(* IEC 61131-3 sources: 2026_Projet_YGO_ExcavatriceDragage/ARCHIVES/Code/PLC_TESTS/BRICKS, 6 files *)

(* ---- FB_TestCheck.st ---- *)
FUNCTION_BLOCK FB_TestCheck
VAR_INPUT
    Config      : ST_TestCheckConfig;
    Evaluate    : BOOL;
END_VAR
VAR_IN_OUT
    ProbeBool   : ARRAY[1..GVL_PLC_Tests_Const.MaxProbeBool] OF BOOL;
    ProbeDint   : ARRAY[1..GVL_PLC_Tests_Const.MaxProbeDint] OF DINT;
    ProbeReal   : ARRAY[1..GVL_PLC_Tests_Const.MaxProbeReal] OF REAL;
END_VAR
VAR_OUTPUT
    Passed       : BOOL;
    Failed       : BOOL;
    Pending      : BOOL;
    FailReason   : E_TestFailReason;
    ObservedBool : BOOL;
    ObservedDint : DINT;
    ObservedReal : REAL;
END_VAR
VAR
    RisingTrig   : R_TRIG;
    FallingTrig  : F_TRIG;
    StableTimer  : TON;
    EvaluateTrig : R_TRIG;
    Cond         : BOOL;
    ProbeIdxLocal : INT;
END_VAR
// === IMPLEMENTATION ===
// Toujours mettre à jour les triggers, avec borne validée AVANT l'accès.
ProbeIdxLocal := Config.ProbeIdx;
IF ProbeIdxLocal >= 1 THEN
    IF ProbeIdxLocal <= GVL_PLC_Tests_Const.MaxProbeBool THEN
        RisingTrig(CLK := ProbeBool[ProbeIdxLocal]);
        FallingTrig(CLK := ProbeBool[ProbeIdxLocal]);
    ELSE
        RisingTrig(CLK := FALSE);
        FallingTrig(CLK := FALSE);
    END_IF;
ELSE
    RisingTrig(CLK := FALSE);
    FallingTrig(CLK := FALSE);
END_IF;

EvaluateTrig(CLK := Evaluate);

IF EvaluateTrig.Q THEN
    Passed := FALSE;
    Failed := FALSE;
    Pending := FALSE;
    FailReason := E_TestFailReason.FAIL_NONE;
    StableTimer(IN := FALSE);
END_IF;

// Mise à jour des valeurs observées
IF Config.ProbeIdx >= 1 THEN
    CASE Config.Kind OF
        E_TestCheckKind.BOOL_EQUAL, E_TestCheckKind.BOOL_RISING, E_TestCheckKind.BOOL_FALLING:
            IF Config.ProbeIdx <= GVL_PLC_Tests_Const.MaxProbeBool THEN
                ObservedBool := ProbeBool[ProbeIdxLocal];
            END_IF;
        E_TestCheckKind.DINT_EQUAL, E_TestCheckKind.DINT_NOT_EQUAL, E_TestCheckKind.DINT_IN_RANGE,
        E_TestCheckKind.WORD_MASK_ALL, E_TestCheckKind.WORD_MASK_ANY, E_TestCheckKind.WORD_MASK_NONE:
            IF Config.ProbeIdx <= GVL_PLC_Tests_Const.MaxProbeDint THEN
                ObservedDint := ProbeDint[ProbeIdxLocal];
            END_IF;
        E_TestCheckKind.REAL_IN_RANGE:
            IF Config.ProbeIdx <= GVL_PLC_Tests_Const.MaxProbeReal THEN
                ObservedReal := ProbeReal[ProbeIdxLocal];
            END_IF;
    END_CASE;
END_IF;

// Évaluation de la condition logique (Cond)
Cond := FALSE;
IF Config.ProbeIdx >= 1 THEN
    CASE Config.Kind OF
        E_TestCheckKind.BOOL_EQUAL:
            IF Config.ProbeIdx <= GVL_PLC_Tests_Const.MaxProbeBool THEN
                Cond := (ObservedBool = Config.ExpectedBool);
            END_IF;

        E_TestCheckKind.BOOL_RISING:
            IF Config.ProbeIdx <= GVL_PLC_Tests_Const.MaxProbeBool THEN
                Cond := RisingTrig.Q;
            END_IF;

        E_TestCheckKind.BOOL_FALLING:
            IF Config.ProbeIdx <= GVL_PLC_Tests_Const.MaxProbeBool THEN
                Cond := FallingTrig.Q;
            END_IF;

        E_TestCheckKind.DINT_EQUAL:
            IF Config.ProbeIdx <= GVL_PLC_Tests_Const.MaxProbeDint THEN
                Cond := (ObservedDint = Config.ExpectedDint);
            END_IF;

        E_TestCheckKind.DINT_NOT_EQUAL:
            IF Config.ProbeIdx <= GVL_PLC_Tests_Const.MaxProbeDint THEN
                Cond := (ObservedDint <> Config.ExpectedDint);
            END_IF;

        E_TestCheckKind.DINT_IN_RANGE:
            IF Config.ProbeIdx <= GVL_PLC_Tests_Const.MaxProbeDint THEN
                Cond := (ObservedDint >= Config.ExpectedMin AND ObservedDint <= Config.ExpectedMax);
            END_IF;

        E_TestCheckKind.WORD_MASK_ALL:
            IF Config.ProbeIdx <= GVL_PLC_Tests_Const.MaxProbeDint THEN
                Cond := ((DINT_TO_WORD(ObservedDint) AND Config.Mask) = Config.Mask);
            END_IF;

        E_TestCheckKind.WORD_MASK_ANY:
            IF Config.ProbeIdx <= GVL_PLC_Tests_Const.MaxProbeDint THEN
                Cond := ((DINT_TO_WORD(ObservedDint) AND Config.Mask) <> 0);
            END_IF;

        E_TestCheckKind.WORD_MASK_NONE:
            IF Config.ProbeIdx <= GVL_PLC_Tests_Const.MaxProbeDint THEN
                Cond := ((DINT_TO_WORD(ObservedDint) AND Config.Mask) = 0);
            END_IF;

        E_TestCheckKind.REAL_IN_RANGE:
            IF Config.ProbeIdx <= GVL_PLC_Tests_Const.MaxProbeReal THEN
                Cond := (ObservedReal >= Config.RealMin AND ObservedReal <= Config.RealMax);
            END_IF;
    END_CASE;
END_IF;

// Application du mode d'évaluation
IF Evaluate THEN
    CASE Config.Mode OF
        E_TestCheckMode.CHECK_INSTANT:
            IF EvaluateTrig.Q THEN
                IF Cond THEN
                    Passed := TRUE;
                    Failed := FALSE;
                    Pending := FALSE;
                ELSE
                    Passed := FALSE;
                    Failed := TRUE;
                    Pending := FALSE;
                    FailReason := E_TestFailReason.FAIL_CHECK;
                END_IF;
            END_IF;

        E_TestCheckMode.CHECK_WAIT_UNTIL:
            IF NOT Passed AND NOT Failed THEN
                StableTimer(IN := Cond, PT := Config.StablePT);
                IF StableTimer.Q THEN
                    Passed := TRUE;
                    Failed := FALSE;
                    Pending := FALSE;
                ELSE
                    Pending := TRUE;
                END_IF;
            END_IF;

        E_TestCheckMode.CHECK_INVARIANT:
            IF NOT Cond THEN
                Passed := FALSE;
                Failed := TRUE;
                Pending := FALSE;
                FailReason := E_TestFailReason.FAIL_INVARIANT;
            ELSE
                Passed := TRUE;
                Failed := FALSE;
                Pending := FALSE;
            END_IF;

        E_TestCheckMode.CHECK_NEVER_DURING:
            IF NOT Failed THEN
                IF Cond THEN
                    Passed := FALSE;
                    Failed := TRUE;
                    Pending := FALSE;
                    FailReason := E_TestFailReason.FAIL_CHECK;
                ELSE
                    Pending := TRUE;
                END_IF;
            END_IF;
    END_CASE;
ELSE
    Passed := FALSE;
    Failed := FALSE;
    Pending := FALSE;
    StableTimer(IN := FALSE);
END_IF;

(* ---- FB_TestEdgeCounter.st ---- *)
FUNCTION_BLOCK FB_TestEdgeCounter
VAR_INPUT
    Arm         : BOOL;
    Signal      : BOOL;
    CountRising : BOOL; // TRUE pour fronts montants, FALSE pour descendants
    ExpectedMin : DINT;
    ExpectedMax : DINT;
END_VAR
VAR_OUTPUT
    Count       : DINT;
    InRange     : BOOL;
END_VAR
VAR
    TrigRising  : R_TRIG;
    TrigFalling : F_TRIG;
END_VAR
// === IMPLEMENTATION ===
TrigRising(CLK := Signal);
TrigFalling(CLK := Signal);

IF NOT Arm THEN
    Count := 0;
    InRange := FALSE;
    RETURN;
END_IF;

IF CountRising AND TrigRising.Q THEN
    Count := Count + 1;
ELSIF NOT CountRising AND TrigFalling.Q THEN
    Count := Count + 1;
END_IF;

InRange := (Count >= ExpectedMin AND Count <= ExpectedMax);

(* ---- FB_TestEventOrder.st ---- *)
FUNCTION_BLOCK FB_TestEventOrder
VAR_INPUT
    Arm       : BOOL;
    EventA    : BOOL;
    EventB    : BOOL;
    TimeoutPT : TIME;
END_VAR
VAR_OUTPUT
    OrderOk   : BOOL;
    Failed    : BOOL;
END_VAR
VAR
    TrigA     : R_TRIG;
    TrigB     : R_TRIG;
    Timer     : TON;
    HasA      : BOOL;
END_VAR
// === IMPLEMENTATION ===
TrigA(CLK := EventA);
TrigB(CLK := EventB);

IF NOT Arm THEN
    OrderOk := FALSE;
    Failed  := FALSE;
    HasA    := FALSE;
    Timer(IN := FALSE);
    RETURN;
END_IF;

// Échec immédiat si B se produit avant A
IF TrigB.Q AND NOT HasA THEN
    Failed  := TRUE;
    OrderOk := FALSE;
END_IF;

// Mémorisation de la survenue de A
IF TrigA.Q AND NOT Failed AND NOT OrderOk THEN
    HasA := TRUE;
END_IF;

// Armement du timeout une fois que A s'est produit
Timer(IN := HasA AND NOT OrderOk AND NOT Failed, PT := TimeoutPT);

IF Timer.Q THEN
    Failed  := TRUE;
    OrderOk := FALSE;
END_IF;

// Validation du succès si B arrive après A et dans les temps
IF HasA AND TrigB.Q AND NOT Failed THEN
    OrderOk := TRUE;
END_IF;

(* ---- FB_TestStimulus.st ---- *)
FUNCTION_BLOCK FB_TestStimulus
VAR_INPUT
    Config     : ST_TestStimAnalogConfig;
    Start      : BOOL;
    Abort      : BOOL;
END_VAR
VAR_OUTPUT
    OutBool    : BOOL;
    OutReal    : REAL;
    OutActive  : BOOL;
    Done       : BOOL;
END_VAR
VAR
    StartTrig   : R_TRIG;
    Timer       : TON;
    SeqTimer    : TON;
    Ramp        : RAMP_REAL;
    ActiveIndex : INT;
    Running     : BOOL;
    Rate        : REAL;
END_VAR
// === IMPLEMENTATION ===
StartTrig(CLK := Start);

// Gestion de l'arrêt ou de l'inactivité
IF Abort OR (NOT Running AND NOT StartTrig.Q) THEN
    Running := FALSE;
    OutActive := FALSE;
    OutBool := FALSE;
    OutReal := 0.0;
    Done := FALSE;
    Timer(IN := FALSE);
    SeqTimer(IN := FALSE);
    Ramp(RESET := TRUE, IN := 0.0);
    RETURN;
END_IF;

// Lancement sur front montant de Start
IF StartTrig.Q THEN
    Running := TRUE;
    Done := FALSE;
    OutActive := TRUE;
    ActiveIndex := 1;
    Timer(IN := FALSE);
    SeqTimer(IN := FALSE);

    CASE Config.Kind OF
        E_TestStimKind.STIM_PULSE_BOOL:
            OutBool := TRUE;
            Timer(IN := TRUE, PT := Config.PulsePT);

        E_TestStimKind.STIM_RAMP_REAL:
            Ramp(RESET := TRUE, IN := Config.StartReal);
            IF Config.RampPT > T#0s THEN
                // Calcul de la vitesse par seconde
                Rate := ABS(Config.TargetReal - Config.StartReal) / (TIME_TO_REAL(Config.RampPT) / 1000.0);
            ELSE
                Rate := ABS(Config.TargetReal - Config.StartReal);
            END_IF;
            Timer(IN := TRUE, PT := Config.RampPT);

        E_TestStimKind.STIM_SEQUENCE_REAL:
            IF Config.SeqCount >= 1 THEN
                OutReal := Config.SeqValues[1];
                SeqTimer(IN := TRUE, PT := Config.SeqDwellPT);
            ELSE
                Running := FALSE;
                OutActive := FALSE;
                Done := TRUE;
            END_IF;
    END_CASE;
END_IF;

// Éxecution logique quand le stimulus tourne
IF Running THEN
    CASE Config.Kind OF
        E_TestStimKind.STIM_PULSE_BOOL:
            Timer();
            IF Timer.Q THEN
                OutBool := FALSE;
                Running := FALSE;
                OutActive := FALSE;
                Done := TRUE;
                Timer(IN := FALSE);
            END_IF;

        E_TestStimKind.STIM_RAMP_REAL:
            Timer();
            Ramp(RESET := FALSE, IN := Config.TargetReal, ASCEND := Rate, DESCEND := Rate, TIMEBASE := T#1s);
            OutReal := Ramp.OUT;
            IF Timer.Q THEN
                OutReal := Config.TargetReal; // Assure la valeur cible exacte à la fin
                Running := FALSE;
                OutActive := FALSE;
                Done := TRUE;
                Timer(IN := FALSE);
            END_IF;

        E_TestStimKind.STIM_SEQUENCE_REAL:
            SeqTimer();
            IF SeqTimer.Q THEN
                SeqTimer(IN := FALSE);
                ActiveIndex := ActiveIndex + 1;
                IF ActiveIndex > Config.SeqCount OR ActiveIndex > GVL_PLC_Tests_Const.MaxSeqValues THEN
                    Running := FALSE;
                    OutActive := FALSE;
                    Done := TRUE;
                ELSE
                    OutReal := Config.SeqValues[ActiveIndex];
                    SeqTimer(IN := TRUE, PT := Config.SeqDwellPT);
                END_IF;
            END_IF;
    END_CASE;
END_IF;

(* ---- FB_TestStopwatch.st ---- *)
FUNCTION_BLOCK FB_TestStopwatch
VAR_INPUT
    Arm             : BOOL;
    StartEvent      : BOOL;
    StopEvent       : BOOL;
    ExpectedMinMs   : DINT;
    ExpectedMaxMs   : DINT;
END_VAR
VAR_OUTPUT
    ElapsedMs       : DINT;
    Done            : BOOL;
    InWindow        : BOOL;
END_VAR
VAR
    StartTrig       : R_TRIG;
    StopTrig        : R_TRIG;
    Running         : BOOL;
    CycleCount      : UDINT;
END_VAR
// === IMPLEMENTATION ===
StartTrig(CLK := StartEvent);
StopTrig(CLK := StopEvent);

IF NOT Arm THEN
    Running := FALSE;
    Done := FALSE;
    InWindow := FALSE;
    ElapsedMs := 0;
    CycleCount := 0;
    RETURN;
END_IF;

IF StartTrig.Q AND NOT Running AND NOT Done THEN
    Running := TRUE;
    CycleCount := 0;
END_IF;

IF Running THEN
    // Incrémente le compteur de cycles
    CycleCount := CycleCount + 1;
    ElapsedMs := UDINT_TO_DINT(CycleCount * INT_TO_UDINT(GVL_PLC_Tests_Const.TaskCycleMs));

    IF StopTrig.Q THEN
        Running := FALSE;
        Done := TRUE;
        InWindow := (ElapsedMs >= ExpectedMinMs AND ElapsedMs <= ExpectedMaxMs);
    END_IF;
END_IF;

(* ---- FB_Timeout.st ---- *)
FUNCTION_BLOCK FB_Timeout
VAR_INPUT
    Active : BOOL;
    PT : TIME;
END_VAR
VAR_OUTPUT
    Elapsed : BOOL;
END_VAR
VAR
    Timer : TON;
END_VAR
// === IMPLEMENTATION ===
Timer(IN := Active, PT := PT);
Elapsed := Timer.Q;
